(*
SPDX-FileCopyrightText: © 2026 Oleksandr Tiutyk <trofimich@gmail.com>
SPDX-License-Identifier: MIT
License: https://opensource.org/license/mit
*)

(*!
<summary>Orders LTIME_OF_DAY values described by generic descriptors.</summary>
<description>
Non-null addresses must reference live LTIME_OF_DAY storage. TypeClass and Size are not validated and no
numeric conversion is performed. Two null addresses compare equal; one null address sorts before a non-null
address. Descriptors are passed by value; payload remains borrowed and is not modified, cloned, released or
retained. IsMemoryOwner does not affect comparison.
</description>
*)

FUNCTION_BLOCK LTimeOfDayComparer EXTENDS TOF_Core.Object IMPLEMENTS TOF_Core.IComparer
VAR_STAT
	//! <summary>Class name shared by all instances of this function block.</summary>
	{attribute 'hide'} 
	_ClassName : STRING := __POUNAME();
END_VAR

{attribute 'monitoring' := 'call'}
PROPERTY ClassName : REFERENCE TO STRING
GET
ClassName REF= _ClassName;
END_GET
END_PROPERTY

(*!
<summary>Compares the first operand with the second using this ordering strategy.</summary>
<description>
Non-null addresses must reference live LTIME_OF_DAY storage. TypeClass and Size are not validated and no
numeric conversion is performed. Two null addresses compare equal; one null address sorts before a non-null
address. Descriptors are passed by value; payload remains borrowed and is not modified, cloned, released or
retained. IsMemoryOwner does not affect comparison. Descendants cannot replace this standard ordering;
implement IComparer separately for a different ordering strategy.
</description>
*)
//!<param name="first">First descriptor; referenced storage is borrowed for the call.</param>
//!<param name="second">Second descriptor; referenced storage is borrowed for the call.</param>
{attribute "object_name" := "Compare"}
METHOD FINAL Compare : TOF_Core.COMPARISON_RESULT
VAR_INPUT
	first : TOF_Core.GENERIC_VALUE;
	second : TOF_Core.GENERIC_VALUE;
END_VAR
VAR
	leftPointer : POINTER TO LTIME_OF_DAY; 
	rightPointer : POINTER TO LTIME_OF_DAY; 
END_VAR
IF first.Address = 0 AND_THEN second.Address = 0 THEN
	Compare := TOF_Core.COMPARISON_RESULT.FIRST_EQUAL_TO_SECOND;
	RETURN;
END_IF

IF first.Address = 0 THEN
	Compare := TOF_Core.COMPARISON_RESULT.FIRST_LESS_THAN_SECOND;
	RETURN;	
END_IF

IF second.Address = 0 THEN
	Compare := TOF_Core.COMPARISON_RESULT.FIRST_GREATER_THAN_SECOND;
	RETURN;	
END_IF

leftPointer := first.Address;
rightPointer := second.Address;

IF leftPointer^ < rightPointer^ THEN
	Compare := TOF_Core.COMPARISON_RESULT.FIRST_LESS_THAN_SECOND;
ELSIF leftPointer^ > rightPointer^ THEN
	Compare := TOF_Core.COMPARISON_RESULT.FIRST_GREATER_THAN_SECOND;
ELSE
	Compare := TOF_Core.COMPARISON_RESULT.FIRST_EQUAL_TO_SECOND;	
END_IF
END_METHOD

{attribute 'monitoring' := 'call'}
PROPERTY NamespaceName : REFERENCE TO STRING
GET
NamespaceName REF= CurrentNamespace.Name;
END_GET
END_PROPERTY

{attribute 'monitoring' := 'call'}
PROPERTY SelfSize : ULINT
GET
SelfSize := XSIZEOF(THIS^);
END_GET
END_PROPERTY

END_FUNCTION_BLOCK

(* stored: Version 1.1.0.1
   POU LTimeOfDayComparer: Id {268f85ac-72d0-4093-81f9-c039f87ef2f8}, SpecialFunc None
   Property ClassName: Id {f7f6ce6a-d55a-4469-8312-391d1993df6b}
   Get Get: Id {88116d14-bc4d-49f1-976c-2d1c84c2989f}
   Method Compare: Id {967550ed-cd5f-4f17-b617-402b2a743ec7}
   Property NamespaceName: Id {0635d7bd-d97a-4f26-9e58-32a637fa3326}
   Get Get: Id {62376183-978d-48d9-9586-104b1886e0c3}
   Property SelfSize: Id {e07ef92b-49ba-4be0-bf90-f7d9d9705a57}
   Get Get: Id {8e9429c6-90a0-45a8-abde-f62672da0a01} *)
